FUNCTION_BLOCK FB_CfcCaller
VAR_OUTPUT
  obReady    : BOOL;
END_VAR
VAR
  fbWorker  : TON;
END_VAR

END_FUNCTION_BLOCK

(* stored: Version 1.1.0.1, ProductVersion 3.1.4024.12
   POU FB_CfcCaller: Id {0a1b2c3d-0000-4000-8000-000000000001}, SpecialFunc None *)
